// TIA Portal V21 export
FUNCTION "FC_AnaWriteInput" : Int   // FC12, SCL
TITLE = Analyzer: write to an input parameter
{ S7_Optimized_Access := 'TRUE' }
// Rule C26f: the input parameter Value is written
// stored: SetENOAutomatically false
   VAR_INPUT
      Value : Int;   // Input value
   END_VAR
BEGIN

       #Value := #Value * 2;
       #FC_AnaWriteInput := #Value;
END_FUNCTION
